(* IEC 61131-3 sources: plcfuzz/testcases/concurrency_candidates, 8 files *)

(* ---- 2333.st ---- *)
PROGRAM helloworld
  VAR
    PB : BOOL;
    LED : BOOL;
  END_VAR

  LED := PB;
END_PROGRAM

CONFIGURATION Config0
  RESOURCE Res0 ON PLC
    TASK task0(INTERVAL := T#20ms,PRIORITY := 0);
    PROGRAM instance0 WITH task0 : helloworld;
  END_RESOURCE
END_CONFIGURATION

(* ---- auto2_new.st ---- *)
TYPE
  LOGLEVEL : (CRITICAL, WARNING, INFO, DEBUG) := INFO;
END_TYPE

PROGRAM program0
   (* Variable definition *)
   VAR
    pb1 AT %IX0.0 : BOOL;
    pb2 AT %IX0.1 : BOOL;
    pb3 AT %IX0.2 : BOOL;
    led AT %QX0.0 : BOOL;
    led2 AT %QX0.1 : BOOL;
    led3 AT %QX0.2 : BOOL;
    led4 AT %QX0.3 : BOOL;
    cstate44 AT %QW1 : INT := 0;
   END_VAR

   (* Control logic *)
CASE cstate44 OF
0:
    IF (( TRUE )) THEN
        cstate44 := 1; led := FALSE; led2 := FALSE; led3 := FALSE; led4 := FALSE;
    END_IF;
1:
    IF ((pb1 = FALSE) AND  ( TRUE ) AND  ( TRUE )) THEN
        cstate44 := 1; led := TRUE; led2 := FALSE; led3 := FALSE; led4 := FALSE;
    ELSIF ((pb1 = TRUE) AND  ( TRUE ) AND  ( TRUE )) THEN
        cstate44 := 3; led := TRUE; led2 := FALSE; led3 := FALSE; led4 := FALSE;
    END_IF;
2:
    IF (( TRUE )) THEN
        cstate44 := 1; led := FALSE; led2 := FALSE; led3 := FALSE; led4 := FALSE;
    END_IF;
3:
    IF ((pb1 = FALSE) AND  ( TRUE ) AND  ( TRUE )) THEN
        cstate44 := 2; led := TRUE; led2 := TRUE; led3 := FALSE; led4 := FALSE;
    ELSIF ((pb1 = TRUE) AND  ( TRUE ) AND  ( TRUE )) THEN
        cstate44 := 4; led := TRUE; led2 := TRUE; led3 := FALSE; led4 := FALSE;
    END_IF;
4:
    IF (( TRUE )) THEN
        cstate44 := 2; led := FALSE; led2 := TRUE; led3 := FALSE; led4 := FALSE;
    END_IF;
END_CASE;

END_PROGRAM

CONFIGURATION Config0
  RESOURCE Res0 ON PLC
    TASK task0(INTERVAL := T#50ms, PRIORITY := 0);
    PROGRAM instance0 WITH task0 : program0;
  END_RESOURCE
END_CONFIGURATION

(* ---- auto_generate.st ---- *)
TYPE
  LOGLEVEL : (CRITICAL, WARNING, INFO, DEBUG) := INFO;
END_TYPE

PROGRAM program0
    VAR_INPUT
        pb1 : BOOL;
    END_VAR
    VAR_OUTPUT
        led : BOOL;
        led2 : BOOL;
    END_VAR
    VAR
        cstate92 : LINT := 0;
    END_VAR

  CASE cstate92 OF
    0:
      IF (TRUE) THEN
        cstate92 := 1;
        led := FALSE;
        led2 := FALSE;
      END_IF;
    1:
      IF (pb1 = FALSE) THEN
        cstate92 := 1;
        led := TRUE;
        led2 := FALSE;
      ELSIF (pb1 = TRUE) THEN
        cstate92 := 2;
        led := TRUE;
        led2 := FALSE;
      END_IF;
    2:
      IF (pb1 = FALSE) THEN
        cstate92 := 3;
        led := TRUE;
        led2 := TRUE;
      ELSIF (pb1 = TRUE) THEN
        cstate92 := 4;
        led := TRUE;
        led2 := TRUE;
      END_IF;
    3:
      IF (TRUE) THEN
        cstate92 := 1;
        led := FALSE;
        led2 := FALSE;
      END_IF;
    4:
      IF (TRUE) THEN
        cstate92 := 3;
        led := FALSE;
        led2 := TRUE;
      END_IF;
  END_CASE;
END_PROGRAM

CONFIGURATION Config0
  VAR_GLOBAL
    PB1 AT %IX0.0 : BOOL;
    LED2 AT %QX0.0 : BOOL;
    LED AT %QX0.1 : BOOL;
  END_VAR
  RESOURCE Res0 ON PLC
    TASK task0(INTERVAL := T#50ms, PRIORITY := 0);
    PROGRAM instance0 WITH task0 : program0;
  END_RESOURCE
END_CONFIGURATION

(* ---- concurrency_candidate.st ---- *)
TYPE
  LOGLEVEL : (CRITICAL, WARNING, INFO, DEBUG) := INFO;
END_TYPE

PROGRAM program0
  VAR
    PB1 AT %IX0.0 : BOOL;
    LED2 AT %QX0.0 : BOOL;
    LED AT %QX0.1 : BOOL;
  END_VAR

  LED2 := LED AND PB1;
  LED := NOT(LED2);
END_PROGRAM

CONFIGURATION Config0

  RESOURCE Res0 ON PLC
    TASK task0(INTERVAL := T#50ms,PRIORITY := 0);
    PROGRAM instance0 WITH task0 : program0;
  END_RESOURCE
END_CONFIGURATION

(* ---- concurrency_test.st ---- *)
TYPE
  LOGLEVEL : (CRITICAL, WARNING, INFO, DEBUG) := INFO;
END_TYPE

PROGRAM program0
  VAR
    PB1 AT %IX0.0 : BOOL;
    LED2 AT %QX0.0 : BOOL;
    LED AT %QX0.1 : BOOL;
  END_VAR

  LED2 := LED AND PB1;
  LED := NOT(LED2);
END_PROGRAM

CONFIGURATION Config0
  RESOURCE Res0 ON PLC
    TASK task0(INTERVAL := T#50ms,PRIORITY := 0);
    PROGRAM instance0 WITH task0 : program0;
  END_RESOURCE
END_CONFIGURATION

(* ---- converted_plc_code.st ---- *)
TYPE
  LOGLEVEL : (CRITICAL, WARNING, INFO, DEBUG) := INFO;
END_TYPE

PROGRAM program0

   (* Variable definition *)
   VAR_INPUT
      pb1	: BOOL;
      pb2	: BOOL;
      pb3	: BOOL;
   END_VAR
   VAR_OUTPUT
      led	: BOOL;
      led2	: BOOL;
      led3	: BOOL;
      led4	: BOOL;
   END_VAR
   VAR
   (* The total number of states equals to 5 *)
      cstate44	: LINT := 0;
   END_VAR

   (* Control logic *)
CASE cstate44 OF
0:
    IF (( TRUE )) THEN
        cstate44 := 1; led := FALSE; led2 := FALSE; led3 := FALSE; led4 := FALSE;
    END_IF;
1:
    IF ((pb1 = FALSE) AND  ( TRUE ) AND  ( TRUE )) THEN
        cstate44 := 1; led := TRUE; led2 := FALSE; led3 := FALSE; led4 := FALSE;
    ELSIF ((pb1 = TRUE) AND  ( TRUE ) AND  ( TRUE )) THEN
        cstate44 := 3; led := TRUE; led2 := FALSE; led3 := FALSE; led4 := FALSE;
    END_IF;
2:
    IF (( TRUE )) THEN
        cstate44 := 1; led := FALSE; led2 := FALSE; led3 := FALSE; led4 := FALSE;
    END_IF;
3:
    IF ((pb1 = FALSE) AND  ( TRUE ) AND  ( TRUE )) THEN
        cstate44 := 2; led := TRUE; led2 := TRUE; led3 := FALSE; led4 := FALSE;
    ELSIF ((pb1 = TRUE) AND  ( TRUE ) AND  ( TRUE )) THEN
        cstate44 := 4; led := TRUE; led2 := TRUE; led3 := FALSE; led4 := FALSE;
    END_IF;
4:
    IF (( TRUE )) THEN
        cstate44 := 2; led := FALSE; led2 := TRUE; led3 := FALSE; led4 := FALSE;
    END_IF;
END_CASE;

END_PROGRAM

CONFIGURATION Config0
  VAR_GLOBAL
    pb1 AT %IX0.0 : BOOL;
    pb2 AT %IX0.1 : BOOL;
    pb3 AT %IX0.2 : BOOL;
    led AT %QX0.0 : BOOL;
    led2 AT %QX0.1 : BOOL;
    led3 AT %QX0.2 : BOOL;
    led4 AT %QX0.3 : BOOL;
  END_VAR
  RESOURCE Res0 ON PLC
    TASK task0(INTERVAL := T#50ms, PRIORITY := 0);
    PROGRAM instance0 WITH task0 : program0;
  END_RESOURCE
END_CONFIGURATION

(* ---- light.st ---- *)
PROGRAM program0
  VAR
    PB1 AT %IX0.0 : BOOL;
    PB2 AT %IX0.1 : BOOL;
    LED AT %QX0.0 : BOOL;
  END_VAR

  LED := NOT(PB2) AND (LED OR PB1);
END_PROGRAM

CONFIGURATION Config0

  RESOURCE Res0 ON PLC
    TASK task0(INTERVAL := T#50ms,PRIORITY := 0);
    PROGRAM instance0 WITH task0 : program0;
  END_RESOURCE
END_CONFIGURATION

(* ---- petrinet_concurrency_example.st ---- *)
TYPE
  LOGLEVEL : (CRITICAL, WARNING, INFO, DEBUG) := INFO;
END_TYPE

PROGRAM program0
  VAR
      IX00 AT %IX0.0 : BOOL;
      IX01 AT %IX0.1 : BOOL;
      IX02 AT %IX0.2 : BOOL;
      IX03 AT %IX0.3 : BOOL;
      IX04 AT %IX0.4 : BOOL;
      QX00 AT %QX0.0 : BOOL;
      QX01 AT %QX0.1 : BOOL;
      QX02 AT %QX0.2 : BOOL;
      QX03 AT %QX0.3 : BOOL;
      QX04 AT %QX0.4 : BOOL;

    END_VAR

    QX04 := QX04 OR IX00 AND NOT IX01;
    QX00 := QX04 AND IX02;
    QX00 := IX04;
    QX01 := QX00 AND IX03;
    QX02 := QX04 AND QX01 AND NOT QX03;
    QX03 := QX04 AND IX02 AND QX02;

END_PROGRAM

CONFIGURATION Config0

  RESOURCE Res0 ON PLC
    TASK task0(INTERVAL := T#50ms,PRIORITY := 0);
    PROGRAM instance0 WITH task0 : program0;
  END_RESOURCE
END_CONFIGURATION
